Fanuc KAREL source: ke00001.compact.KL

PROGRAM KE00001
%STACKSIZE=65535
%PRIORITY=65535
%NOLOCKGROUP
%ENVIRONMENT REGOPE
VAR
I : INTEGER
S : STRING[80]
STATUS : INTEGER
BEGIN
I=1
GET_PREG_CMT(I,S,STATUS)
END KE00001
